// TIA Portal V20 export
Screen "190FX3LhSliderFixtureLayout"  1276x673
  ScreenItem "Line_Header_X0_Y64" at 0,64 size 1276x0  Type=HmiLine
  ScreenItem "permanentareaborderrectangle" at 0,0 size 0x0  Type=HmiRectangle
  ScreenItem "Button_Back" at 2,2 size 90x60  Type=HmiButton
  ScreenItem "Move_Legend" at 1182,2 size 90x60  Type=HmiButton
  ScreenItem "Fusszeile_Button_ManualOPMode1_2" at 279,2 size 90x60  Type=HmiButton
  ScreenItem "文本域_22" at 1126,369 size 104x23  Type=HmiTextBox
  ScreenItem "Fusszeile_Button_ManualOPMode1_1" at 95,2 size 90x60  Type=HmiButton
  ScreenItem "Fusszeile_Button_ManualOPMode1_3" at 187,2 size 90x60  Type=HmiButton
  ScreenItem "Fusszeile_Button_ManualOPMode1_4" at 997,2 size 90x60  Type=HmiButton
  ScreenItem "Fusszeile_Button_ManualOPMode1_5" at 902,1 size 90x60  Type=HmiButton
  ScreenItem "文本域_14" at 936,-172 size 140x40  Type=HmiTextBox
  ScreenItem "Title_ScreenOverview_X390_Y2_1" at 384,5 size 510x57  Type=HmiTextBox
  ScreenItem "Graphic view_1" at 260,212 size 560x296  Type=HmiGraphicView
  ScreenItem "文本域_5" at -1,82 size 120x40  Type=HmiTextBox
  ScreenItem "文本域_27" at -1,126 size 120x40  Type=HmiTextBox
  ScreenItem "面板容器_22" at 1063,402 size 96x32  Type=HmiFaceplateContainer
  ScreenItem "面板容器_23" at 1173,402 size 96x32  Type=HmiFaceplateContainer
  ScreenItem "文本域_21" at 679,90 size 140x40  Type=HmiTextBox
  ScreenItem "Line_4" at 609,241 size 255x25  Type=HmiLine
  ScreenItem "Faceplate container_6" at 889,249 size 59x45  Type=HmiFaceplateContainer
  ScreenItem "文本域_12" at 869,209 size 100x40  Type=HmiTextBox
  ScreenItem "Line_1" at 532,174 size 150x98  Type=HmiLine
  ScreenItem "文本域_6" at 73,206 size 140x40  Type=HmiTextBox
  ScreenItem "面板容器_1" at 80,247 size 144x51  Type=HmiFaceplateContainer
  ScreenItem "Line_2" at 220,239 size 194x50  Type=HmiLine
  ScreenItem "文本域_7" at 236,90 size 100x40  Type=HmiTextBox
  ScreenItem "Line_3" at 294,180 size 128x81  Type=HmiLine
  ScreenItem "文本域_8" at 95,356 size 100x40  Type=HmiTextBox
  ScreenItem "Faceplate container_2" at 115,399 size 59x45  Type=HmiFaceplateContainer
  ScreenItem "Line_5" at 198,301 size 241x66  Type=HmiLine
  ScreenItem "文本域_9" at 410,516 size 100x40  Type=HmiTextBox
  ScreenItem "Faceplate container_3" at 430,556 size 59x45  Type=HmiFaceplateContainer
  ScreenItem "Line_6" at 466,344 size 22x172  Type=HmiLine
  ScreenItem "文本域_10" at 869,373 size 100x40  Type=HmiTextBox
  ScreenItem "Faceplate container_4" at 889,413 size 59x45  Type=HmiFaceplateContainer
  ScreenItem "Line_7" at 607,299 size 258x90  Type=HmiLine
  ScreenItem "文本域_13" at 456,90 size 140x40  Type=HmiTextBox
  ScreenItem "Line_9" at 510,159 size 10x128  Type=HmiLine
  ScreenItem "文本域_15" at 564,516 size 100x40  Type=HmiTextBox
  ScreenItem "Faceplate container_5" at 584,556 size 59x45  Type=HmiFaceplateContainer
  ScreenItem "Line_10" at 555,341 size 33x171  Type=HmiLine
  ScreenItem "LSicar_Valve8Pos_LeftHomeRightWork_WithPB_2" at 1099,271 size 160x53  Type=HmiFaceplateContainer
  ScreenItem "文本域_2" at 1094,246 size 165x23  Type=HmiTextBox
  ScreenItem "LSicar_Valve8Pos_LeftHomeRightWork_WithPB_1" at 1099,183 size 160x53  Type=HmiFaceplateContainer
  ScreenItem "文本域_1" at 1099,160 size 156x23  Type=HmiTextBox
  ScreenItem "LSicar_Valve8Pos_LeftHomeRightWork_WithPB_5" at 1099,95 size 160x53  Type=HmiFaceplateContainer
  ScreenItem "文本域_3" at 1107,71 size 139x22  Type=HmiTextBox
  ScreenItem "面板容器_8" at 682,136 size 144x51  Type=HmiFaceplateContainer
  ScreenItem "面板容器_4" at 459,136 size 144x51  Type=HmiFaceplateContainer
  ScreenItem "Faceplate container_1" at 256,136 size 59x45  Type=HmiFaceplateContainer
  ScreenItem "面板容器_2" at 1090,4 size 88x58  Type=HmiFaceplateContainer
  ScreenItem "OPMode1_Blocked" at 1164,6 size 14x14  Type=HmiGraphicView
  ScreenItem "OPMode4_Foreground_Blocked" at 1089,2 size 88x58  Type=HmiGraphicView
